FUNCTION_BLOCK Conveyor (* CAT Function Block Type *)
  (* Standard: 61499-2 *)
  (* Version 0.0, 11/22/2026, Schneider Electric, Conveyor CAT with 4 belt outputs and 6 lightweight StopPoints *)
  PACKAGE Main;
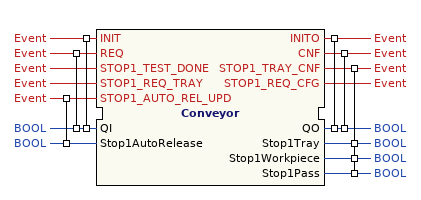
  EVENT_INPUT
    INIT WITH QI; (* Initialization Request *)
    REQ WITH QI; (* Normal Execution Request *)
    STOP1_TEST_DONE; (* Primary Station 1 Testing pass-complete notification for Stop 1 *)
    STOP1_REQ_TRAY; (* Request current Station 1 tray and workpiece sensor states *)
    STOP1_AUTO_REL_UPD WITH Stop1AutoRelease; (* Update Stop 1 automatic release enable from Station 1 *)
  END_EVENT
  EVENT_OUTPUT
    INITO WITH QO; (* Initialization Confirm *)
    CNF WITH QO; (* Execution Confirmation *)
    STOP1_TRAY_CNF WITH Stop1Tray, Stop1Workpiece, Stop1Pass; (* Station 1 tray and workpiece sensor update *)
    STOP1_REQ_CFG; (* Request initial Stop 1 auto-release configuration from Testing on startup *)
  END_EVENT
  VAR_INPUT
    QI : BOOL := TRUE; (* Input event qualifier *)
    Stop1AutoRelease : BOOL := FALSE; (* Stop 1 automatic release enable (Auto S1 AND Auto-Rel) *)
  END_VAR
  VAR_OUTPUT
    QO : BOOL; (* Output event qualifier *)
    Stop1Tray : BOOL; (* Tray present at Stop 1 (Station 1) *)
    Stop1Workpiece : BOOL; (* Workpiece present on tray at Stop 1 (Station 1) *)
    Stop1Pass : BOOL; (* Stopper 1 pass-through or releasing state (TRUE=Down, FALSE=Up/Blocking) *)
  END_VAR
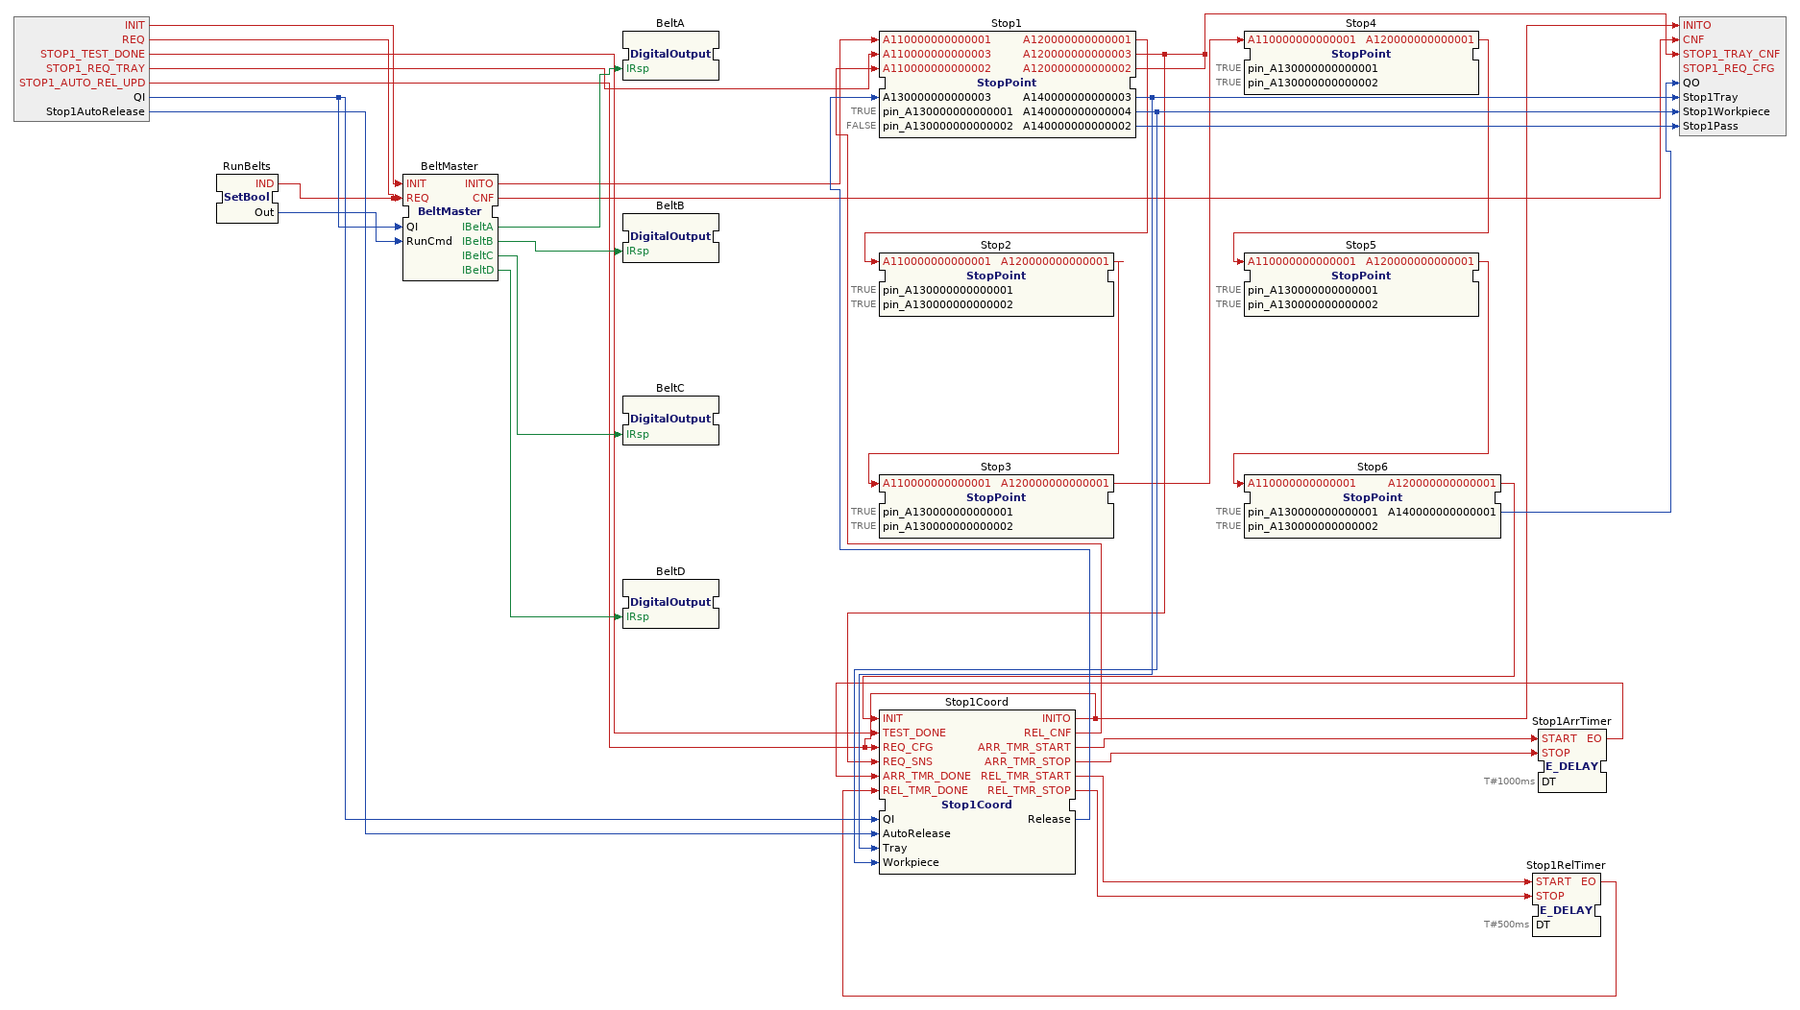
  FBS
    BeltA : DigitalOutput;
    BeltB : DigitalOutput;
    BeltC : DigitalOutput;
    BeltD : DigitalOutput;
    RunBelts : SetBool;
    BeltMaster : BeltMaster;
    Stop1 : StopPoint(pin_A130000000000001 := TRUE, pin_A130000000000002 := FALSE);
    Stop2 : StopPoint(pin_A130000000000001 := TRUE, pin_A130000000000002 := TRUE);
    Stop3 : StopPoint(pin_A130000000000001 := TRUE, pin_A130000000000002 := TRUE);
    Stop4 : StopPoint(pin_A130000000000001 := TRUE, pin_A130000000000002 := TRUE);
    Stop5 : StopPoint(pin_A130000000000001 := TRUE, pin_A130000000000002 := TRUE);
    Stop6 : StopPoint(pin_A130000000000001 := TRUE, pin_A130000000000002 := TRUE);
    Stop1Coord : Stop1Coord;
    Stop1ArrTimer : E_DELAY(DT := T#1000ms);
    Stop1RelTimer : E_DELAY(DT := T#500ms);
  END_FBS
  EVENT_CONNECTIONS
    INIT TO BeltMaster.INIT;
    BeltMaster.INITO TO Stop1.A110000000000001;
    Stop1.A120000000000001 TO Stop2.A110000000000001;
    Stop2.A120000000000001 TO Stop3.A110000000000001;
    Stop3.A120000000000001 TO Stop4.A110000000000001;
    Stop4.A120000000000001 TO Stop5.A110000000000001;
    Stop5.A120000000000001 TO Stop6.A110000000000001;
    Stop6.A120000000000001 TO Stop1Coord.INIT;
    Stop1Coord.INITO TO INITO;
    RunBelts.IND TO BeltMaster.REQ;
    REQ TO BeltMaster.REQ;
    BeltMaster.CNF TO CNF;
    STOP1_TEST_DONE TO Stop1Coord.TEST_DONE;
    STOP1_AUTO_REL_UPD TO Stop1Coord.REQ_CFG;
    STOP1_REQ_TRAY TO Stop1.A110000000000003;
    Stop1.A120000000000003 TO STOP1_TRAY_CNF;
    Stop1.A120000000000003 TO Stop1Coord.REQ_SNS;
    Stop1.A120000000000002 TO STOP1_TRAY_CNF;
    Stop1Coord.REL_CNF TO Stop1.A110000000000002;
    Stop1Coord.ARR_TMR_START TO Stop1ArrTimer.START;
    Stop1Coord.ARR_TMR_STOP TO Stop1ArrTimer.STOP;
    Stop1ArrTimer.EO TO Stop1Coord.ARR_TMR_DONE;
    Stop1Coord.REL_TMR_START TO Stop1RelTimer.START;
    Stop1Coord.REL_TMR_STOP TO Stop1RelTimer.STOP;
    Stop1RelTimer.EO TO Stop1Coord.REL_TMR_DONE;
    Stop1Coord.INITO TO Stop1Coord.REQ_CFG;
  END_CONNECTIONS
  DATA_CONNECTIONS
    QI TO BeltMaster.QI;
    QI TO Stop1Coord.QI;
    RunBelts.Out TO BeltMaster.RunCmd;
    Stop6.A140000000000001 TO QO;
    Stop1AutoRelease TO Stop1Coord.AutoRelease;
    Stop1.A140000000000003 TO Stop1Coord.Tray;
    Stop1.A140000000000004 TO Stop1Coord.Workpiece;
    Stop1Coord.Release TO Stop1.A130000000000003;
    Stop1.A140000000000003 TO Stop1Tray;
    Stop1.A140000000000004 TO Stop1Workpiece;
    Stop1.A140000000000002 TO Stop1Pass;
  END_CONNECTIONS
  ADAPTER_CONNECTIONS
    BeltMaster.IBeltA TO BeltA.IRsp;
    BeltMaster.IBeltB TO BeltB.IRsp;
    BeltMaster.IBeltC TO BeltC.IRsp;
    BeltMaster.IBeltD TO BeltD.IRsp;
  END_CONNECTIONS
END_FUNCTION_BLOCK
